Fanuc KAREL source: KD00045.KL

PROGRAM KD00045
%NOLOCKGROUP
%DEFGROUP = 1
VAR
  I: INTEGER
  J: INTEGER
  B: BOOLEAN
  R: REAL
  S: STRING[80]
  P: POSITION
BEGIN
  MOVE TO P
END KD00045
